(* PLC project Vn_move, Beckhoff Automation GmbH TwinCAT PLC Control 3.5.13.21 *)
(* stored: creationDateTime 1970-01-01T00:00:00 *)

PROGRAM Vn_move

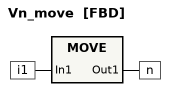
(* FBD diagram, written out as Structured Text *)
n := i1;
END_PROGRAM
